// TIA Portal V20 export
Screen "OrderManagement"  1276x673
  ScreenItem "permanentareaborderrectangle" at 0,0 size 0x0  Type=HmiRectangle
  ScreenItem "Button_Back" at 2,2 size 90x44  Type=HmiButton
  ScreenItem "线_1" at 0,46 size 1363x0  Type=HmiLine
  ScreenItem "Title_OPMode1_ScreenOverview_X390_Y2" at 418,5 size 500x30  Type=HmiTextBox
  ScreenItem "Faceplate container_1" at 2,70 size 1273x555  Type=HmiFaceplateContainer
